FUNCTION_BLOCK Test (* Composite Function Block Type *)
  (* Standard: 61499-2 *)
  (* Version 0.0, 7/14/2016, Andrei, nxtControl GmbH, template *)
  PACKAGE Main;
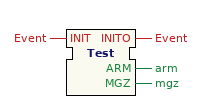
  EVENT_INPUT
    INIT; (* Initialization Request *)
  END_EVENT
  EVENT_OUTPUT
    INITO; (* Initialization Confirm *)
  END_EVENT
  PLUGS
    ARM : arm;
    MGZ : mgz;
  END_PLUGS
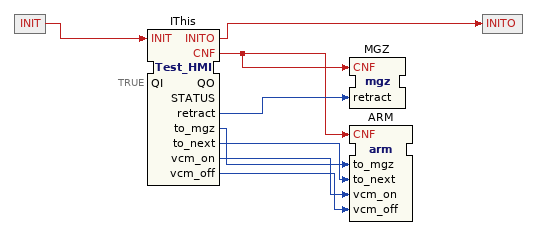
  FBS
    IThis : Test_HMI(QI := TRUE);
  END_FBS
  EVENT_CONNECTIONS
    INIT TO IThis.INIT;
    IThis.INITO TO INITO;
    IThis.CNF TO MGZ.CNF;
    IThis.CNF TO ARM.CNF;
  END_CONNECTIONS
  DATA_CONNECTIONS
    IThis.retract TO MGZ.retract;
    IThis.to_mgz TO ARM.to_mgz;
    IThis.to_next TO ARM.to_next;
    IThis.vcm_on TO ARM.vcm_on;
    IThis.vcm_off TO ARM.vcm_off;
  END_CONNECTIONS
END_FUNCTION_BLOCK
